(* IEC 61131-3 sources: iolistgen/pytests/golden/gen_fixture/src/GVLs/Generated, 6 files *)

(* ---- GVL_CfgProject.gvl.st ---- *)
// AUTO-GENERATED by iolistgen 0.2.0 — не редактировать; источник: gen_fixture.csv
// SHA-256 перечня 3ace79e7a28b; генератор st-codesys
// Назначение: уставки проекта — Cfg устройств из перечня сигналов, те же инициализаторы, что у GVL_Persist.
// PRG_ApplyProjectCfg копирует их в GVL_Persist (контракт plc-process-lib 18.3, правило 2).
{attribute 'qualified_only'}
VAR_GLOBAL CONSTANT
    // --- dev_no 1: LT201 — Уровень в резервуаре чистой воды (AnalogInput) ---
    // lint:allow STL007 структура-константа: имя как у GVL_Persist.stLT201Cfg (контракт 18.3, правило 2)
    stLT201Cfg : PL.ST_AnalogInputCfg := (
        rRangeHi_eu := 4.0,
        tFilter := T#2S,
        astLimit := [
            (xEnable := TRUE, rSetpoint_eu := 3.6, tOnDelay := T#2S, tOffDelay := T#1S),  // 0 HH
            (xEnable := TRUE, rSetpoint_eu := 3.2, rHyst_eu := 0.05, tOnDelay := T#2S, tOffDelay := T#1S),  // 1 H
            (xEnable := TRUE, rSetpoint_eu := 0.8, tOnDelay := T#2S, tOffDelay := T#1S),  // 2 L
            (xEnable := TRUE, rSetpoint_eu := 0.4, tOnDelay := T#2S, tOffDelay := T#1S)  // 3 LL
        ],
        udiAlarmIdBase := 10,
        astAlarm := [
            (ePriority := PL.E_AlarmPriority.High),  // 0 HH
            (ePriority := PL.E_AlarmPriority.Medium),  // 1 H
            (ePriority := PL.E_AlarmPriority.Medium),  // 2 L
            (ePriority := PL.E_AlarmPriority.High),  // 3 LL
            (ePriority := PL.E_AlarmPriority.Medium),  // 4 Failure
            (ePriority := PL.E_AlarmPriority.Low),  // 5 OutOfRange
            (ePriority := PL.E_AlarmPriority.None),  // 6 (резерв)
            (ePriority := PL.E_AlarmPriority.None)  // 7 (резерв)
        ]
    );
    // --- dev_no 2: PT201 — Давление на всасе (AnalogInput) ---
    // lint:allow STL007 структура-константа: имя как у GVL_Persist.stPT201Cfg (контракт 18.3, правило 2)
    stPT201Cfg : PL.ST_AnalogInputCfg := (
        eInput := PL.E_AiInputType.Raw,
        rRangeHi_eu := 16.0,
        rRawHi_cnt := 16000.0,
        astLimit := [
            (xEnable := FALSE),  // 0 HH
            (xEnable := FALSE),  // 1 H
            (xEnable := TRUE, rSetpoint_eu := 1.0),  // 2 L
            (xEnable := FALSE)  // 3 LL
        ],
        udiAlarmIdBase := 20,
        astAlarm := [
            (ePriority := PL.E_AlarmPriority.Medium),  // 0 HH
            (ePriority := PL.E_AlarmPriority.Low),  // 1 H
            (ePriority := PL.E_AlarmPriority.Low),  // 2 L
            (ePriority := PL.E_AlarmPriority.Medium),  // 3 LL
            (ePriority := PL.E_AlarmPriority.Medium),  // 4 Failure
            (ePriority := PL.E_AlarmPriority.Low),  // 5 OutOfRange
            (ePriority := PL.E_AlarmPriority.None),  // 6 (резерв)
            (ePriority := PL.E_AlarmPriority.None)  // 7 (резерв)
        ]
    );
    // --- dev_no 3: TE201 — Температура воды (AnalogInput) ---
    // lint:allow STL007 структура-константа: имя как у GVL_Persist.stTE201Cfg (контракт 18.3, правило 2)
    stTE201Cfg : PL.ST_AnalogInputCfg := (
        eInput := PL.E_AiInputType.Norm01,
        rRangeLo_eu := -50.0,
        rRangeHi_eu := 150.0,
        astLimit := [
            (xEnable := FALSE),  // 0 HH
            (xEnable := TRUE, rSetpoint_eu := 80.0),  // 1 H
            (xEnable := FALSE),  // 2 L
            (xEnable := FALSE)  // 3 LL
        ],
        udiAlarmIdBase := 30
    );
    // --- dev_no 4: LS201 — Поплавок «перелив» (DigitalInput) ---
    // lint:allow STL007 структура-константа: имя как у GVL_Persist.stLS201Cfg (контракт 18.3, правило 2)
    stLS201Cfg : PL.ST_DigitalInputCfg := (
        xInvert := TRUE,
        tOnDelay := T#2S,
        udiAlarmIdBase := 40,
        astAlarm := [
            (ePriority := PL.E_AlarmPriority.High),  // 0 State
            (ePriority := PL.E_AlarmPriority.Medium),  // 1 Failure
            (ePriority := PL.E_AlarmPriority.None),  // 2 (резерв)
            (ePriority := PL.E_AlarmPriority.None),  // 3 (резерв)
            (ePriority := PL.E_AlarmPriority.None),  // 4 (резерв)
            (ePriority := PL.E_AlarmPriority.None),  // 5 (резерв)
            (ePriority := PL.E_AlarmPriority.None),  // 6 (резерв)
            (ePriority := PL.E_AlarmPriority.None)  // 7 (резерв)
        ]
    );
    // --- dev_no 5: ES201 — Кнопка аварийного останова на щите (DigitalInput) ---
    // lint:allow STL007 структура-константа: имя как у GVL_Persist.stES201Cfg (контракт 18.3, правило 2)
    stES201Cfg : PL.ST_DigitalInputCfg := (
        udiAlarmIdBase := 50,
        astAlarm := [
            (ePriority := PL.E_AlarmPriority.Critical),  // 0 State
            (ePriority := PL.E_AlarmPriority.Medium),  // 1 Failure
            (ePriority := PL.E_AlarmPriority.None),  // 2 (резерв)
            (ePriority := PL.E_AlarmPriority.None),  // 3 (резерв)
            (ePriority := PL.E_AlarmPriority.None),  // 4 (резерв)
            (ePriority := PL.E_AlarmPriority.None),  // 5 (резерв)
            (ePriority := PL.E_AlarmPriority.None),  // 6 (резерв)
            (ePriority := PL.E_AlarmPriority.None)  // 7 (резерв)
        ]
    );
    // --- dev_no 6: PWR2 — Напряжение на секции шин (DigitalInput) ---
    // lint:allow STL007 структура-константа: имя как у GVL_Persist.stPWR2Cfg (контракт 18.3, правило 2)
    stPWR2Cfg : PL.ST_DigitalInputCfg := (
        xAlarmOnTrue := FALSE,
        udiAlarmIdBase := 60,
        astAlarm := [
            (ePriority := PL.E_AlarmPriority.High),  // 0 State
            (ePriority := PL.E_AlarmPriority.Medium),  // 1 Failure
            (ePriority := PL.E_AlarmPriority.None),  // 2 (резерв)
            (ePriority := PL.E_AlarmPriority.None),  // 3 (резерв)
            (ePriority := PL.E_AlarmPriority.None),  // 4 (резерв)
            (ePriority := PL.E_AlarmPriority.None),  // 5 (резерв)
            (ePriority := PL.E_AlarmPriority.None),  // 6 (резерв)
            (ePriority := PL.E_AlarmPriority.None)  // 7 (резерв)
        ]
    );
    // --- dev_no 11: M201 — Насос промывки (Motor) ---
    // lint:allow STL007 структура-константа: имя как у GVL_Persist.stM201Cfg (контракт 18.3, правило 2)
    stM201Cfg : PL.ST_MotorCfg := (tFbStart := T#3S, tFbStop := T#8S, tMinStop := T#20S, udiAlarmIdBase := 110);
    // --- dev_no 12: P201 — Насос Н1 (MotorVfd) ---
    // lint:allow STL007 структура-константа: имя как у GVL_Persist.stP201Cfg (контракт 18.3, правило 2)
    stP201Cfg : PL.ST_MotorCfg := (uiMaxStartsPerHour := 6, stVfd := (rSpeedMin_pct := 25.0), udiAlarmIdBase := 120);
    // --- dev_no 13: P202 — Насос Н2 (MotorVfd) ---
    // lint:allow STL007 структура-константа: имя как у GVL_Persist.stP202Cfg (контракт 18.3, правило 2)
    stP202Cfg : PL.ST_MotorCfg := (stVfd := (xFbFromComm := FALSE, xCommLossIsFault := FALSE), udiAlarmIdBase := 130);
    // --- dev_no 21: FV201 — Задвижка на напоре (Valve) ---
    // lint:allow STL007 структура-константа: имя как у GVL_Persist.stFV201Cfg (контракт 18.3, правило 2)
    stFV201Cfg : PL.ST_ValveCfg := (
        tTravel := T#1M15S,
        xTorqueUsed := TRUE,
        xCloseOnTorque := TRUE,
        udiAlarmIdBase := 210
    );
    // --- dev_no 22: XV201 — Клапан сброса (Valve) ---
    // lint:allow STL007 структура-константа: имя как у GVL_Persist.stXV201Cfg (контракт 18.3, правило 2)
    stXV201Cfg : PL.ST_ValveCfg := (
        eType := PL.E_ValveType.SolenoidEtc,
        xZsoUsed := FALSE,
        eSafePos := PL.E_ValveSafePos.Open,
        udiAlarmIdBase := 220
    );
    // --- dev_no 31: FCV201 — Клапан рециркуляции (ControlValve) ---
    // lint:allow STL007 структура-константа: имя как у GVL_Persist.stFCV201Cfg (контракт 18.3, правило 2)
    stFCV201Cfg : PL.ST_ControlValveCfg := (
        rSafePos_pct := 100.0,
        eFaultAction := PL.E_CvFaultAction.SafePos,
        xFbUsed := TRUE,
        tDev := T#40S,
        udiAlarmIdBase := 310
    );
    // --- dev_no 32: ZT201 — Клапан рециркуляции: положение (AnalogInput) ---
    // lint:allow STL007 структура-константа: имя как у GVL_Persist.stZT201Cfg (контракт 18.3, правило 2)
    stZT201Cfg : PL.ST_AnalogInputCfg := (udiAlarmIdBase := 320);
    // --- dev_no 41: LIC201 — Регулятор уровня в резервуаре чистой воды (Pid) ---
    // lint:allow STL007 структура-константа: имя как у GVL_Persist.stLIC201Cfg (контракт 18.3, правило 2)
    stLIC201Cfg : PL.ST_PidCfg := (
        eAction := PL.E_PidAction.Direct,
        rKp := 2.0,
        rTi_s := 120.0,
        rPvMax_eu := 4.0,
        rSpMin_eu := 0.5,
        rSpMax_eu := 3.5,
        xUseOutAct := TRUE,
        udiAlarmIdBase := 410,
        astAlarm := [
            (ePriority := PL.E_AlarmPriority.Low),  // 0 PvInvalid
            (ePriority := PL.E_AlarmPriority.None),  // 1 (резерв)
            (ePriority := PL.E_AlarmPriority.None),  // 2 (резерв)
            (ePriority := PL.E_AlarmPriority.None),  // 3 (резерв)
            (ePriority := PL.E_AlarmPriority.None),  // 4 (резерв)
            (ePriority := PL.E_AlarmPriority.None),  // 5 (резерв)
            (ePriority := PL.E_AlarmPriority.None),  // 6 (резерв)
            (ePriority := PL.E_AlarmPriority.None)  // 7 (резерв)
        ]
    );
END_VAR

(* ---- GVL_Devices.gvl.st ---- *)
// AUTO-GENERATED by iolistgen 0.2.0 — не редактировать; источник: gen_fixture.csv
// SHA-256 перечня 3ace79e7a28b; генератор st-codesys
// Назначение: экземпляры устройств plc-process-lib (объявление без параметров, контракт 20). Логика станции пишет их
// входы автоматики и читает выходы; HMI и SCADA читают stSts.
{attribute 'qualified_only'}
VAR_GLOBAL
    fbLT201 : PL.FB_AnalogInput;  // 1 · Уровень в резервуаре чистой воды
    fbPT201 : PL.FB_AnalogInput;  // 2 · Давление на всасе
    fbTE201 : PL.FB_AnalogInput;  // 3 · Температура воды
    fbLS201 : PL.FB_DigitalInput;  // 4 · Поплавок «перелив»
    fbES201 : PL.FB_DigitalInput;  // 5 · Кнопка аварийного останова на щите
    fbPWR2 : PL.FB_DigitalInput;  // 6 · Напряжение на секции шин
    fbM201 : PL.FB_Motor;  // 11 · Насос промывки
    fbP201 : PL.FB_MotorVfd;  // 12 · Насос Н1
    fbP202 : PL.FB_MotorVfd;  // 13 · Насос Н2
    fbFV201 : PL.FB_Valve;  // 21 · Задвижка на напоре
    fbXV201 : PL.FB_Valve;  // 22 · Клапан сброса
    fbFCV201 : PL.FB_ControlValve;  // 31 · Клапан рециркуляции
    fbZT201 : PL.FB_AnalogInput;  // 32 · Клапан рециркуляции: положение
    fbLIC201 : PL.FB_PID;  // 41 · Регулятор уровня в резервуаре чистой воды
END_VAR

(* ---- GVL_DevIdx.gvl.st ---- *)
// AUTO-GENERATED by iolistgen 0.2.0 — не редактировать; источник: gen_fixture.csv
// SHA-256 перечня 3ace79e7a28b; генератор st-codesys
// Назначение: номера устройств dev_no (контракт plc-process-lib 20.1): тревоги устройства — dev_no · 10 + слот; для
// SCADA и логики станции.
{attribute 'qualified_only'}
VAR_GLOBAL CONSTANT
    LT201 : UINT := 1;  // AnalogInput · Уровень в резервуаре чистой воды
    PT201 : UINT := 2;  // AnalogInput · Давление на всасе
    TE201 : UINT := 3;  // AnalogInput · Температура воды
    LS201 : UINT := 4;  // DigitalInput · Поплавок «перелив»
    ES201 : UINT := 5;  // DigitalInput · Кнопка аварийного останова на щите
    PWR2 : UINT := 6;  // DigitalInput · Напряжение на секции шин
    M201 : UINT := 11;  // Motor · Насос промывки
    P201 : UINT := 12;  // MotorVfd · Насос Н1
    P202 : UINT := 13;  // MotorVfd · Насос Н2
    FV201 : UINT := 21;  // Valve · Задвижка на напоре
    XV201 : UINT := 22;  // Valve · Клапан сброса
    FCV201 : UINT := 31;  // ControlValve · Клапан рециркуляции
    ZT201 : UINT := 32;  // AnalogInput · Клапан рециркуляции: положение
    LIC201 : UINT := 41;  // Pid · Регулятор уровня в резервуаре чистой воды
END_VAR

(* ---- GVL_Hmi.gvl.st ---- *)
// AUTO-GENERATED by iolistgen 0.2.0 — не редактировать; источник: gen_fixture.csv
// SHA-256 перечня 3ace79e7a28b; генератор st-codesys
// Назначение: команды HMI и SCADA устройствам (ST_<Dev>Cmd, контракт plc-process-lib 1 и 2.1). WebVisu и OPC UA пишут
// сюда напрямую; команды по Modbus — только через адаптер приложения (импульс по фронту).
{attribute 'qualified_only'}
VAR_GLOBAL
    xApplyProjectCfg : BOOL;  // импульс: применить уставки проекта (PRG_ApplyProjectCfg); сбрасывает PRG_Devices
    stLT201Cmd : PL.ST_AnalogInputCmd;  // 1 · Уровень в резервуаре чистой воды
    stPT201Cmd : PL.ST_AnalogInputCmd;  // 2 · Давление на всасе
    stTE201Cmd : PL.ST_AnalogInputCmd;  // 3 · Температура воды
    stLS201Cmd : PL.ST_DigitalInputCmd;  // 4 · Поплавок «перелив»
    stES201Cmd : PL.ST_DigitalInputCmd;  // 5 · Кнопка аварийного останова на щите
    stPWR2Cmd : PL.ST_DigitalInputCmd;  // 6 · Напряжение на секции шин
    stM201Cmd : PL.ST_MotorCmd;  // 11 · Насос промывки
    stP201Cmd : PL.ST_MotorCmd;  // 12 · Насос Н1
    stP202Cmd : PL.ST_MotorCmd;  // 13 · Насос Н2
    stFV201Cmd : PL.ST_ValveCmd;  // 21 · Задвижка на напоре
    stXV201Cmd : PL.ST_ValveCmd;  // 22 · Клапан сброса
    stFCV201Cmd : PL.ST_ControlValveCmd;  // 31 · Клапан рециркуляции
    stZT201Cmd : PL.ST_AnalogInputCmd;  // 32 · Клапан рециркуляции: положение
    stLIC201Cmd : PL.ST_PidCmd;  // 41 · Регулятор уровня в резервуаре чистой воды
END_VAR

(* ---- GVL_IO.gvl.st ---- *)
// AUTO-GENERATED by iolistgen 0.2.0 — не редактировать; источник: gen_fixture.csv
// SHA-256 перечня 3ace79e7a28b; генератор st-codesys
// Назначение: переменные ввода-вывода перечня сигналов — каналы модулей, обмен Modbus, адаптеры ПЧ. Адресов %I/%Q в
// коде нет: каналы привязываются в дереве устройств (I/O Mapping → «Map to existing variable»), значения Modbus пишет и
// читает слой Modbus, переменные ПЧ — адаптеры приложения (docs/MANUAL_STEPS.md).
{attribute 'qualified_only'}
VAR_GLOBAL
    // === Входы модулей ввода-вывода (DI, AI): дерево устройств, I/O Mapping → Map to existing variable ===
    rLT201_mA : REAL;  // A1.1 · LT201 · Уровень в резервуаре чистой воды · 0…4 м
    rTE201 : REAL;  // A1.2 · TE201 · Температура воды · -50…150 °C
    rP202_ACT : REAL;  // A1.3 · P202_ACT · Насос Н2: выход частоты 4–20 мА · 0…50 Гц · адаптер ПЧ
    rZT201_mA : REAL;  // A1.4 · ZT201 · Клапан рециркуляции: положение · 0…100 %
    xLT201_CHF : BOOL;  // D1.1 · LT201_CHF · Уровень в резервуаре: отказ канала модуля
    xLS201 : BOOL;  // D1.2 · LS201 · Поплавок «перелив»
    xLS201_CHF : BOOL;  // D1.3 · LS201_CHF · Поплавок «перелив»: обрыв цепи
    xPWR2 : BOOL;  // D1.4 · PWR2 · Напряжение на секции шин
    xM201_FB : BOOL;  // D1.5 · M201_FB · Насос промывки: в работе
    xM201_FLT : BOOL;  // D1.6 · M201_FLT · Насос промывки: авария УПП
    xM201_LOC : BOOL;  // D1.7 · M201_LOC · Насос промывки: режим «Местное»
    xP201_FLT : BOOL;  // D1.8 · P201_FLT · Насос Н1: тепловое реле
    xP201_LOC : BOOL;  // D1.9 · P201_LOC · Насос Н1: режим «Местное»
    xP202_FB : BOOL;  // D1.10 · P202_FB · Насос Н2: реле «работа» ПЧ
    xFV201_ZSO : BOOL;  // D2.1 · FV201_ZSO · Задвижка на напоре: открыта
    xFV201_ZSC : BOOL;  // D2.2 · FV201_ZSC · Задвижка на напоре: закрыта
    xFV201_TQO : BOOL;  // D2.3 · FV201_TQO · Задвижка на напоре: муфта открытия
    xFV201_TQC : BOOL;  // D2.4 · FV201_TQC · Задвижка на напоре: муфта закрытия
    xFV201_FLT : BOOL;  // D2.5 · FV201_FLT · Задвижка на напоре: авария привода
    xFV201_LOC : BOOL;  // D2.6 · FV201_LOC · Задвижка на напоре: «Местное»
    xXV201_ZSC : BOOL;  // D2.7 · XV201_ZSC · Клапан сброса: закрыт
    xFCV201_POSF : BOOL;  // D2.8 · FCV201_POSF · Клапан рециркуляции: авария позиционера
    xFCV201_LOC : BOOL;  // D2.9 · FCV201_LOC · Клапан рециркуляции: позиционер в местном

    // === Выходы модулей ввода-вывода (DO, AO): дерево устройств, I/O Mapping → Map to existing variable ===
    rP202_REF : REAL;  // A2.1 · P202_REF · Насос Н2: задание частоты 4–20 мА · 0…50 Гц · адаптер ПЧ
    rFCV201_OUT_mA : REAL;  // A2.2 · FCV201_OUT · Клапан рециркуляции: задание положения · 0…100 %
    // A2.3 · LIC201_SPI · Регулятор уровня: задание на индикатор щита · 0…4 м · без ФБ — код приложения
    rLIC201_SPI : REAL;
    xM201_RUN : BOOL;  // Q1.1 · M201_RUN · Насос промывки: команда «Работа»
    xM201_RST : BOOL;  // Q1.2 · M201_RST · Насос промывки: сброс аварии УПП
    xP202_RUN : BOOL;  // Q1.3 · P202_RUN · Насос Н2: команда «Работа»
    xFV201_OPN : BOOL;  // Q1.4 · FV201_OPN · Задвижка на напоре: открыть
    xFV201_CLS : BOOL;  // Q1.5 · FV201_CLS · Задвижка на напоре: закрыть
    xXV201 : BOOL;  // Q1.6 · XV201 · Клапан сброса

    // === Modbus, ПЛК — master, чтение: значения пишет слой Modbus ===
    wP201_STW : WORD;  // RS485-1 · слейв 1 · FC3 4x 10 WORD · P201_STW · Насос Н1: слово состояния ПЧ · адаптер ПЧ
    // RS485-1 · слейв 1 · FC3 4x 12 REAL HL · P201_ACT · Насос Н1: фактическая частота · 0…50 Гц · адаптер ПЧ
    rP201_ACT : REAL;
    wP202_STW : WORD;  // RS485-1 · слейв 2 · FC3 4x 10 WORD · P202_STW · Насос Н2: слово состояния ПЧ · адаптер ПЧ
    iPT201 : INT;  // RS485-1 · слейв 5 · FC4 3x 10 INT · PT201 · Давление на всасе · 0…16 бар
    xES201 : BOOL;  // RS485-1 · слейв 7 · FC2 1x 0 BOOL · ES201 · Кнопка аварийного останова на щите

    // === Modbus, ПЛК — master, запись: значения читает слой Modbus ===
    wP201_CTW : WORD;  // RS485-1 · слейв 1 · FC6 4x 0 WORD · P201_CTW · Насос Н1: слово управления ПЧ · адаптер ПЧ
    // RS485-1 · слейв 1 · FC16 4x 2 REAL HL · P201_REF · Насос Н1: задание частоты · 0…50 Гц · адаптер ПЧ
    rP201_REF : REAL;

    // === Состояние обмена со слейвами: пишет слой Modbus (TRUE — обмен исправен) ===
    xMbOk_RS485_1_S1 : BOOL;  // линия RS485-1, слейв 1: обмен исправен
    xMbOk_RS485_1_S2 : BOOL;  // линия RS485-1, слейв 2: обмен исправен
    xMbOk_RS485_1_S5 : BOOL;  // линия RS485-1, слейв 5: обмен исправен
    xMbOk_RS485_1_S7 : BOOL;  // линия RS485-1, слейв 7: обмен исправен

    // === Адаптеры ПЧ (код приложения) → ФБ: разобранное слово состояния и фактическая скорость ===
    xP201_CommOk : BOOL;  // P201: обмен с ПЧ исправен → xCommOk
    xP201_VfdRun : BOOL;  // P201: ПЧ в работе (слово состояния) → xVfdRunning
    xP201_VfdReady : BOOL;  // P201: ПЧ готов к пуску (слово состояния) → xVfdReady
    xP201_VfdFault : BOOL;  // P201: авария ПЧ (слово состояния) → xVfdFault
    rP201_SpeedAct_pct : REAL;  // P201: фактическая скорость, % → rSpeedAct_pct
    xP202_CommOk : BOOL;  // P202: обмен с ПЧ исправен → xCommOk
    xP202_VfdRun : BOOL;  // P202: ПЧ в работе (слово состояния) → xVfdRunning
    xP202_VfdReady : BOOL;  // P202: ПЧ готов к пуску (слово состояния) → xVfdReady
    xP202_VfdFault : BOOL;  // P202: авария ПЧ (слово состояния) → xVfdFault
    rP202_SpeedAct_pct : REAL;  // P202: фактическая скорость, % → rSpeedAct_pct

    // === ФБ → адаптеры ПЧ: задание скорости и команды для слова управления ===
    rP201_SpeedRef_pct : REAL;  // P201: задание на ПЧ, % ← rSpeedRef_pct
    xP201_VfdQRun : BOOL;  // P201: команда «работа» для слова управления ← xQRun
    xP201_VfdQReset : BOOL;  // P201: импульс сброса аварии ПЧ для слова управления ← xQReset
    rP202_SpeedRef_pct : REAL;  // P202: задание на ПЧ, % ← rSpeedRef_pct
END_VAR

(* ---- GVL_Persist.pvl.st ---- *)
// AUTO-GENERATED by iolistgen 0.2.0 — не редактировать; источник: gen_fixture.csv
// SHA-256 перечня 3ace79e7a28b; генератор st-codesys
// Назначение: объект Persistent Variables (контракт plc-process-lib 18.3): Cfg и Retain устройств, по переменной на
// устройство, по возрастанию dev_no. Новое устройство — dev_no больше прежних (переменные встают в конец); типы
// существующих переменных не меняются. Начальные значения — уставки перечня; после загрузки действуют сохранённые
// значения, уставки проекта применяет PRG_ApplyProjectCfg. Объект создаётся в CODESYS вручную (docs/MANUAL_STEPS.md);
// «Reorder List and Clear Gaps» не выполнять.
VAR_GLOBAL PERSISTENT RETAIN
    uiLayoutVersion : UINT := 1;  // версия раскладки списка
    // --- dev_no 1: LT201 — Уровень в резервуаре чистой воды (AnalogInput, без Retain) ---
    stLT201Cfg : PL.ST_AnalogInputCfg := (
        rRangeHi_eu := 4.0,
        tFilter := T#2S,
        astLimit := [
            (xEnable := TRUE, rSetpoint_eu := 3.6, tOnDelay := T#2S, tOffDelay := T#1S),  // 0 HH
            (xEnable := TRUE, rSetpoint_eu := 3.2, rHyst_eu := 0.05, tOnDelay := T#2S, tOffDelay := T#1S),  // 1 H
            (xEnable := TRUE, rSetpoint_eu := 0.8, tOnDelay := T#2S, tOffDelay := T#1S),  // 2 L
            (xEnable := TRUE, rSetpoint_eu := 0.4, tOnDelay := T#2S, tOffDelay := T#1S)  // 3 LL
        ],
        udiAlarmIdBase := 10,
        astAlarm := [
            (ePriority := PL.E_AlarmPriority.High),  // 0 HH
            (ePriority := PL.E_AlarmPriority.Medium),  // 1 H
            (ePriority := PL.E_AlarmPriority.Medium),  // 2 L
            (ePriority := PL.E_AlarmPriority.High),  // 3 LL
            (ePriority := PL.E_AlarmPriority.Medium),  // 4 Failure
            (ePriority := PL.E_AlarmPriority.Low),  // 5 OutOfRange
            (ePriority := PL.E_AlarmPriority.None),  // 6 (резерв)
            (ePriority := PL.E_AlarmPriority.None)  // 7 (резерв)
        ]
    );
    // --- dev_no 2: PT201 — Давление на всасе (AnalogInput, без Retain) ---
    stPT201Cfg : PL.ST_AnalogInputCfg := (
        eInput := PL.E_AiInputType.Raw,
        rRangeHi_eu := 16.0,
        rRawHi_cnt := 16000.0,
        astLimit := [
            (xEnable := FALSE),  // 0 HH
            (xEnable := FALSE),  // 1 H
            (xEnable := TRUE, rSetpoint_eu := 1.0),  // 2 L
            (xEnable := FALSE)  // 3 LL
        ],
        udiAlarmIdBase := 20,
        astAlarm := [
            (ePriority := PL.E_AlarmPriority.Medium),  // 0 HH
            (ePriority := PL.E_AlarmPriority.Low),  // 1 H
            (ePriority := PL.E_AlarmPriority.Low),  // 2 L
            (ePriority := PL.E_AlarmPriority.Medium),  // 3 LL
            (ePriority := PL.E_AlarmPriority.Medium),  // 4 Failure
            (ePriority := PL.E_AlarmPriority.Low),  // 5 OutOfRange
            (ePriority := PL.E_AlarmPriority.None),  // 6 (резерв)
            (ePriority := PL.E_AlarmPriority.None)  // 7 (резерв)
        ]
    );
    // --- dev_no 3: TE201 — Температура воды (AnalogInput, без Retain) ---
    stTE201Cfg : PL.ST_AnalogInputCfg := (
        eInput := PL.E_AiInputType.Norm01,
        rRangeLo_eu := -50.0,
        rRangeHi_eu := 150.0,
        astLimit := [
            (xEnable := FALSE),  // 0 HH
            (xEnable := TRUE, rSetpoint_eu := 80.0),  // 1 H
            (xEnable := FALSE),  // 2 L
            (xEnable := FALSE)  // 3 LL
        ],
        udiAlarmIdBase := 30
    );
    // --- dev_no 4: LS201 — Поплавок «перелив» (DigitalInput, без Retain) ---
    stLS201Cfg : PL.ST_DigitalInputCfg := (
        xInvert := TRUE,
        tOnDelay := T#2S,
        udiAlarmIdBase := 40,
        astAlarm := [
            (ePriority := PL.E_AlarmPriority.High),  // 0 State
            (ePriority := PL.E_AlarmPriority.Medium),  // 1 Failure
            (ePriority := PL.E_AlarmPriority.None),  // 2 (резерв)
            (ePriority := PL.E_AlarmPriority.None),  // 3 (резерв)
            (ePriority := PL.E_AlarmPriority.None),  // 4 (резерв)
            (ePriority := PL.E_AlarmPriority.None),  // 5 (резерв)
            (ePriority := PL.E_AlarmPriority.None),  // 6 (резерв)
            (ePriority := PL.E_AlarmPriority.None)  // 7 (резерв)
        ]
    );
    // --- dev_no 5: ES201 — Кнопка аварийного останова на щите (DigitalInput, без Retain) ---
    stES201Cfg : PL.ST_DigitalInputCfg := (
        udiAlarmIdBase := 50,
        astAlarm := [
            (ePriority := PL.E_AlarmPriority.Critical),  // 0 State
            (ePriority := PL.E_AlarmPriority.Medium),  // 1 Failure
            (ePriority := PL.E_AlarmPriority.None),  // 2 (резерв)
            (ePriority := PL.E_AlarmPriority.None),  // 3 (резерв)
            (ePriority := PL.E_AlarmPriority.None),  // 4 (резерв)
            (ePriority := PL.E_AlarmPriority.None),  // 5 (резерв)
            (ePriority := PL.E_AlarmPriority.None),  // 6 (резерв)
            (ePriority := PL.E_AlarmPriority.None)  // 7 (резерв)
        ]
    );
    // --- dev_no 6: PWR2 — Напряжение на секции шин (DigitalInput, без Retain) ---
    stPWR2Cfg : PL.ST_DigitalInputCfg := (
        xAlarmOnTrue := FALSE,
        udiAlarmIdBase := 60,
        astAlarm := [
            (ePriority := PL.E_AlarmPriority.High),  // 0 State
            (ePriority := PL.E_AlarmPriority.Medium),  // 1 Failure
            (ePriority := PL.E_AlarmPriority.None),  // 2 (резерв)
            (ePriority := PL.E_AlarmPriority.None),  // 3 (резерв)
            (ePriority := PL.E_AlarmPriority.None),  // 4 (резерв)
            (ePriority := PL.E_AlarmPriority.None),  // 5 (резерв)
            (ePriority := PL.E_AlarmPriority.None),  // 6 (резерв)
            (ePriority := PL.E_AlarmPriority.None)  // 7 (резерв)
        ]
    );
    // --- dev_no 11: M201 — Насос промывки (Motor) ---
    stM201Cfg : PL.ST_MotorCfg := (tFbStart := T#3S, tFbStop := T#8S, tMinStop := T#20S, udiAlarmIdBase := 110);
    stM201Retain : PL.ST_DeviceRetain;  // режим, вывод из работы, наработка, операции
    // --- dev_no 12: P201 — Насос Н1 (MotorVfd) ---
    stP201Cfg : PL.ST_MotorCfg := (uiMaxStartsPerHour := 6, stVfd := (rSpeedMin_pct := 25.0), udiAlarmIdBase := 120);
    stP201Retain : PL.ST_DeviceRetain;  // режим, вывод из работы, наработка, операции
    // --- dev_no 13: P202 — Насос Н2 (MotorVfd) ---
    stP202Cfg : PL.ST_MotorCfg := (stVfd := (xFbFromComm := FALSE, xCommLossIsFault := FALSE), udiAlarmIdBase := 130);
    stP202Retain : PL.ST_DeviceRetain;  // режим, вывод из работы, наработка, операции
    // --- dev_no 21: FV201 — Задвижка на напоре (Valve) ---
    stFV201Cfg : PL.ST_ValveCfg := (
        tTravel := T#1M15S,
        xTorqueUsed := TRUE,
        xCloseOnTorque := TRUE,
        udiAlarmIdBase := 210
    );
    stFV201Retain : PL.ST_DeviceRetain;  // режим, вывод из работы, наработка, операции
    // --- dev_no 22: XV201 — Клапан сброса (Valve) ---
    stXV201Cfg : PL.ST_ValveCfg := (
        eType := PL.E_ValveType.SolenoidEtc,
        xZsoUsed := FALSE,
        eSafePos := PL.E_ValveSafePos.Open,
        udiAlarmIdBase := 220
    );
    stXV201Retain : PL.ST_DeviceRetain;  // режим, вывод из работы, наработка, операции
    // --- dev_no 31: FCV201 — Клапан рециркуляции (ControlValve) ---
    stFCV201Cfg : PL.ST_ControlValveCfg := (
        rSafePos_pct := 100.0,
        eFaultAction := PL.E_CvFaultAction.SafePos,
        xFbUsed := TRUE,
        tDev := T#40S,
        udiAlarmIdBase := 310
    );
    stFCV201Retain : PL.ST_DeviceRetain;  // режим, вывод из работы, наработка, операции
    // --- dev_no 32: ZT201 — Клапан рециркуляции: положение (AnalogInput, без Retain) ---
    stZT201Cfg : PL.ST_AnalogInputCfg := (udiAlarmIdBase := 320);
    // --- dev_no 41: LIC201 — Регулятор уровня в резервуаре чистой воды (Pid) ---
    stLIC201Cfg : PL.ST_PidCfg := (
        eAction := PL.E_PidAction.Direct,
        rKp := 2.0,
        rTi_s := 120.0,
        rPvMax_eu := 4.0,
        rSpMin_eu := 0.5,
        rSpMax_eu := 3.5,
        xUseOutAct := TRUE,
        udiAlarmIdBase := 410,
        astAlarm := [
            (ePriority := PL.E_AlarmPriority.Low),  // 0 PvInvalid
            (ePriority := PL.E_AlarmPriority.None),  // 1 (резерв)
            (ePriority := PL.E_AlarmPriority.None),  // 2 (резерв)
            (ePriority := PL.E_AlarmPriority.None),  // 3 (резерв)
            (ePriority := PL.E_AlarmPriority.None),  // 4 (резерв)
            (ePriority := PL.E_AlarmPriority.None),  // 5 (резерв)
            (ePriority := PL.E_AlarmPriority.None),  // 6 (резерв)
            (ePriority := PL.E_AlarmPriority.None)  // 7 (резерв)
        ]
    );
    stLIC201Retain : PL.ST_DeviceRetain;  // режим, вывод из работы, наработка, операции
END_VAR
